{region 'Documentation'}
(*!
<summary>Checks inequality with the forbidden USINT value.</summary>
*)
{endregion}
FUNCTION_BLOCK AssertNotEqual_USInt EXTENDS AssertionBase
VAR_INPUT
    IN : USINT; //! Actual value checked or observed by this Assertion.
    Expected : USINT; //! Value that must differ from IN under this Assertion's comparison rules.
END_VAR

SUPER^();

{region 'Documentation'}
(*!
<summary>Check inequality with the forbidden USINT value.</summary>
*)
{endregion}
METHOD PROTECTED Assert
VAR
    Message : STRING(GVL_Constants.MessageLength);
    ExpectedText : STRING(GVL_Constants.AssertionValueLength);
    ActualText : STRING(GVL_Constants.AssertionValueLength);
END_VAR
IF NOT EvaluationActive THEN
    RETURN;
END_IF;

IF Result = E_Result.Error THEN
    RETURN;
END_IF;

IF Result = E_Result.Failed THEN
    RETURN;
END_IF;

IF IN = Expected THEN
    ExpectedText := USINT_TO_STRING(Expected);
    ActualText := USINT_TO_STRING(IN);
    Message := CONCAT('Assertion failed: values are equal but should differ. NotExpected = ',
        ExpectedText);
    Message := CONCAT(Message, ', Actual = ');
    Message := CONCAT(Message, ActualText);
    Message := CONCAT(Message, '.');
    Fail(Message := Message);
    RETURN;
END_IF;

Pass();
END_METHOD

END_FUNCTION_BLOCK

(* stored: Version 1.1.0.1
   POU AssertNotEqual_USInt: Id {a3b4d2ba-05b4-43cc-b3e9-3ffd8973da60}, SpecialFunc None
   Folder Internal: Id {9efd27d7-b945-4b6d-9393-fd1dab5306aa}
   Method Assert: Id {a1a59a2d-01d1-4568-898a-03e6b4cdabfe} *)
